Fanuc KAREL source: KO00122.KL

PROGRAM KO00122
%NOLOCKGROUP
VAR
  A: ARRAY[2] OF SHORT
  B: INTEGER
  OUT: REAL
BEGIN
  A[1] = 1
  B = 2
  OUT = ATAN2(A[1], B)
END KO00122
